FUNCTION_BLOCK FB_Location_Workshop
VAR_INPUT
    stInputs : ST_HomeInputs;
END_VAR

VAR_IN_OUT
    stOutputs : ST_HomeOutputs;
END_VAR

VAR
    nMainHandle : UINT := 0;
    fbMainButton : FB_Button;
    fbMainLight : FB_Light;
END_VAR

IF nMainHandle = 0 OR nMainHandle > GVL_HomeLimits.cMaxLights THEN
    RETURN;
END_IF

fbMainButton(
    bPressed := stInputs.aButtons[GVL_WorkshopConfig.stMainLight.nButtonIndex]
);

fbMainLight(
    bToggle := fbMainButton.bShortPress,
    bSetValid := stInputs.aLightCommands[nMainHandle].bValid AND NOT fbMainButton.bShortPress,
    bSetOn := stInputs.aLightCommands[nMainHandle].bOn
);

stOutputs.aLights[nMainHandle].bValid := TRUE;
stOutputs.aLights[nMainHandle].bOn := fbMainLight.bOn;

METHOD PUBLIC RegisterLights : BOOL
VAR_IN_OUT
    fbCatalog : FB_LightCatalog;
END_VAR
nMainHandle := fbCatalog.RegisterLight(stDefinition := GVL_WorkshopConfig.stMainLight);
RegisterLights := nMainHandle <> 0;
END_METHOD

END_FUNCTION_BLOCK

(* stored: Version 1.1.0.1
   POU FB_Location_Workshop: Id {ec750405-3890-4654-994f-cda0aa9720a1}, SpecialFunc None
   Method RegisterLights: Id {f80a87d0-80a4-45ea-a3db-c5a6ceca75b7} *)
